(* IEC 61131-3 sources: llm-plc-st-eval/data/definitivo/claude-sonnet-4-6/B7/zero_shot, 3 files *)

(* ---- ejec_1.st ---- *)
```pascal
// Selección de fuente de mando de bomba
// Sin memoria entre ciclos → FUNCTION (salida puramente combinacional)

FUNCTION SelBomba : BOOL
VAR_INPUT
    modoAuto  : BOOL; // TRUE = modo automático, FALSE = modo manual
    btnManual : BOOL; // Botón de mando en modo manual
    nivelBajo : BOOL; // Señal de nivel bajo (activa = nivel bajo detectado)
END_VAR

// En modo automático la bomba sigue a nivelBajo;
// en modo manual la bomba sigue a btnManual.
SelBomba := (modoAuto AND nivelBajo) OR (NOT modoAuto AND btnManual);

END_FUNCTION
```

(* ---- ejec_2.st ---- *)
```pascal
// Selección de fuente de mando de una bomba.
// Sin memoria entre ciclos: la salida depende solo de las entradas actuales.
FUNCTION SelBomba : BOOL
    VAR_INPUT
        modoAuto  : BOOL; // TRUE = modo automático, FALSE = modo manual
        btnManual : BOOL; // Botón de mando en modo manual
        nivelBajo : BOOL; // Señal de nivel bajo (activa = nivel bajo detectado)
    END_VAR

    // En modo automático la bomba arranca por nivel bajo;
    // en modo manual obedece directamente al botón.
    IF modoAuto THEN
        SelBomba := nivelBajo;  // Modo automático: manda el nivel
    ELSE
        SelBomba := btnManual;  // Modo manual: manda el botón
    END_IF;

END_FUNCTION
```

(* ---- ejec_3.st ---- *)
```pascal
// Selección de fuente de mando para una bomba.
// Sin memoria entre ciclos: la salida depende solo de las entradas actuales.
FUNCTION SelBomba : BOOL
    VAR_INPUT
        modoAuto  : BOOL; // TRUE = modo automático, FALSE = modo manual
        btnManual : BOOL; // Botón de mando en modo manual
        nivelBajo : BOOL; // Señal de nivel bajo (activa la bomba en modo auto)
    END_VAR

    // En modo automático la bomba sigue a nivelBajo;
    // en modo manual la bomba sigue al botón.
    IF modoAuto THEN
        SelBomba := nivelBajo;
    ELSE
        SelBomba := btnManual;
    END_IF;

END_FUNCTION
```
